SUBAPPLICATION INI_IN_AND_STORE_AR2_OVERRIDE (* Wie INI_IN_AND_STORE_AR2, aber MIT Override-Moeglichkeit: Socket OVERRIDE_ACTIVE (AX) erzwingt bei TRUE kontinuierlich einen konfigurierten Wert (Parameter INIT_VAL an LIT_Override, Default 0.0) statt des Live-VT-Werts. Bei OVERRIDE_ACTIVE=FALSE (unbenutzt) identisches Verhalten wie INI_IN_AND_STORE_AR2. *)
  (* Standard: 61499-2; Description: Copyright (c) 2026 Meisterschulen am Ostbahnhof This program and the accompanying materials are made available under the terms of the Eclipse Public License 2.0 which is available at https://www.eclipse.org/legal/epl-2.0/ SPDX-License-Identifier: EPL-2.0 *)
  (* Version 1.0, 2026-10-13, Franz Höpfinger, Meisterschulen am Ostbahnhof, AR2-Pendant zu INI_IN_AND_STORE_AUDI2_OVERRIDE: NumericValue_PHYSA + SEL_Override (AR_AX_SEL_AR, G=OVERRIDE_ACTIVE) + AR_TO_AR2 + INI_AR2, AR_TO_AR2.AR_OUT gesplittet auf Q_NumericValue_PHYSA (VT-Anzeige) und VALUEO (weiterer Consumer). Im Unterschied zu AUDI2 (Enum/Dropdown, 1=Deaktiviert) ist AR ein kontinuierlicher physikalischer Wert - der Override-Wert hat hier keine feste Business-Bedeutung, sondern ist ueber INIT_VAL an LIT_Override frei konfigurierbar (Default 0.0). *)
  PACKAGE MyLib::sys;
  IMPORT isobus::UT::Q::const::IDs::ID_NULL;
  IMPORT logiBUS::utils::conversion::phys::NumericObjectPool_S;
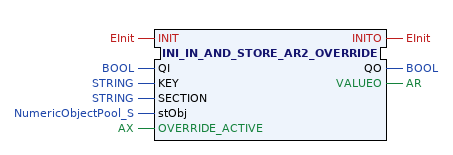
  EVENT_INPUT
    INIT : EInit; (* Initialization Request *)
  END_EVENT
  EVENT_OUTPUT
    INITO : EInit; (* Initialization Confirm *)
  END_EVENT
  VAR_INPUT
    QI : BOOL := TRUE; (* Quality Input - TRUE to enable service *)
    KEY : STRING; (* Key name. *)
    SECTION : STRING; (* Section name. *)
    stObj : logiBUS::utils::conversion::phys::NumericObjectPool_S := (u16ObjId := ID_NULL, r32Scale := 1.0, i32Offset := 0, u8Decimals := 0);
  END_VAR
  VAR_OUTPUT
    QO : BOOL; (* Quality Output - TRUE if service executed successfully *)
  END_VAR
  SOCKETS
    OVERRIDE_ACTIVE : adapter::types::unidirectional::AX; (* Kontinuierlich TRUE erzwingt den ueber LIT_Override.INIT_VAL konfigurierten Wert, unabhaengig vom Live-VT-Wert. FALSE (unbenutzt, Default bei den meisten Aufrufern) = unveraendertes Verhalten. *)
  END_SOCKETS
  PLUGS
    VALUEO : adapter::types::unidirectional::AR;
  END_PLUGS
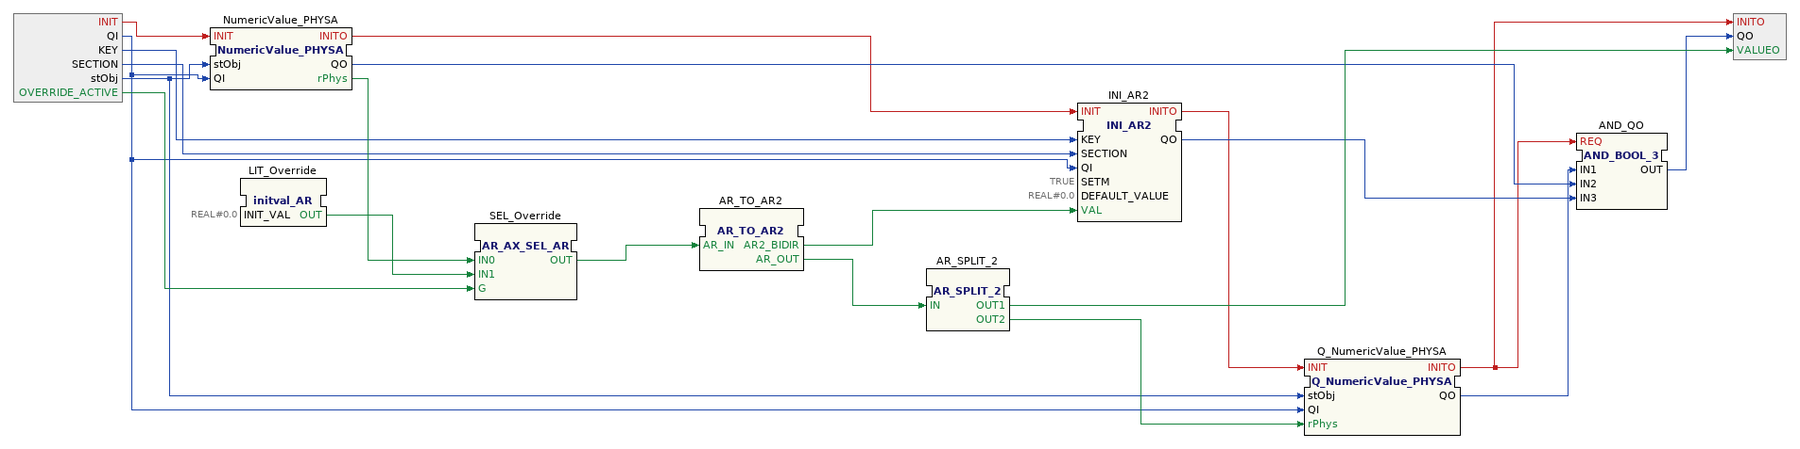
  (* SETM=TRUE - der Boot-Wert laedt so oder so automatisch (INIT -> INITO -> GET -> GETO, unabhaengig von SETM). SETM=TRUE sorgt dafuer, dass auch eine LIVE-Aenderung waehrend des laufenden Betriebs sofort bestaetigt/zurueckgemeldet wird - wichtig, falls der frische Wert noch im selben Lauf weiterverwendet werden soll (z.B. hier ueber VALUEO). *)
  FBS
    NumericValue_PHYSA : isobus::UT::io::NumericValue::NumericValue_PHYSA;
    LIT_Override : adapter::types::unidirectional::AR::initval::initval_AR(INIT_VAL := REAL#0.0); (* Override-Wert, per Parameter konfigurierbar *)
    SEL_Override : adapter::iec61131::selection::AR_AX_SEL_AR; (* IN0=Live-VT-Wert (unveraendert), IN1=Override-Wert, G=OVERRIDE_ACTIVE *)
    AR_TO_AR2 : adapter::conversion::bidirectional::AR_TO_AR2;
    INI_AR2 : eclipse4diac::storage::INI_AR2(SETM := TRUE, DEFAULT_VALUE := REAL#0.0);
    AR_SPLIT_2 : adapter::events::unidirectional::AR_SPLIT_2;
    Q_NumericValue_PHYSA : isobus::UT::Q::Q_NumericValue_PHYSA;
    AND_QO : iec61131::booleanOperators::AND_BOOL_3;
  END_FBS
  EVENT_CONNECTIONS
    INIT TO NumericValue_PHYSA.INIT;
    NumericValue_PHYSA.INITO TO INI_AR2.INIT;
    INI_AR2.INITO TO Q_NumericValue_PHYSA.INIT;
    Q_NumericValue_PHYSA.INITO TO INITO;
    Q_NumericValue_PHYSA.INITO TO AND_QO.REQ;
  END_CONNECTIONS
  DATA_CONNECTIONS
    stObj TO Q_NumericValue_PHYSA.stObj;
    KEY TO INI_AR2.KEY;
    SECTION TO INI_AR2.SECTION;
    stObj TO NumericValue_PHYSA.stObj;
    QI TO Q_NumericValue_PHYSA.QI;
    QI TO NumericValue_PHYSA.QI;
    QI TO INI_AR2.QI;
    Q_NumericValue_PHYSA.QO TO AND_QO.IN1;
    NumericValue_PHYSA.QO TO AND_QO.IN2;
    INI_AR2.QO TO AND_QO.IN3;
    AND_QO.OUT TO QO;
  END_CONNECTIONS
  ADAPTER_CONNECTIONS
    NumericValue_PHYSA.rPhys TO SEL_Override.IN0;
    LIT_Override.OUT TO SEL_Override.IN1;
    OVERRIDE_ACTIVE TO SEL_Override.G;
    SEL_Override.OUT TO AR_TO_AR2.AR_IN;
    AR_TO_AR2.AR2_BIDIR TO INI_AR2.VAL;
    AR_TO_AR2.AR_OUT TO AR_SPLIT_2.IN;
    AR_SPLIT_2.OUT1 TO VALUEO;
    AR_SPLIT_2.OUT2 TO Q_NumericValue_PHYSA.rPhys;
  END_CONNECTIONS
END_SUBAPPLICATION
